(* PLC project c.project, CODESYS CODESYS V3.5 SP17 Patch 3 *)
(* stored: creationDateTime 2026-10-19T00:00:00, modificationDateTime 2026-10-19T00:00:00 *)

FUNCTION_BLOCK FB_L
VAR_INPUT
    a : BOOL;
    b : BOOL;
END_VAR
VAR_OUTPUT
    q : BOOL;
    r : BOOL;
END_VAR

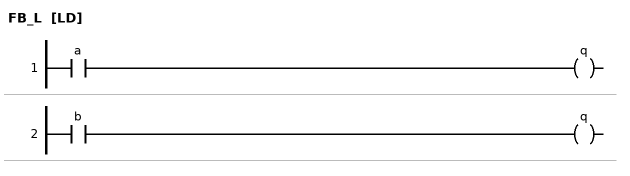
(* LD diagram, written out as Structured Text *)

q := a;

q := b;
END_FUNCTION_BLOCK
